// TIA Portal V21 export
// export: Created 2026-11-21T12:56:43.079897Z, ExportSetting WithDefaults, DisplayName Totally Integrated Automation Portal, DisplayVersion V21, DisplayName STEP 7 Professional, DisplayVersion V21, DisplayName STEP 7 Safety, DisplayVersion V21, DisplayName Tech WebApplication, DisplayVersion V21, DisplayName WinCC Basic/Comfort/Advanced, DisplayVersion V21, DisplayName WinCC Unified, DisplayVersion V21
VAR_GLOBAL   // PLC tag table "IO"
   Start_Line AT %I10.0 : Bool;   // First input of DI_Main
   Lamp_Line AT %Q0.0 : Bool;   // First output of DQ_Main
END_VAR
